(* IEC 61131-3 sources: 2026_Projet_YGO_ExcavatriceDragage/CODE/J_SUPERVISION/_TYPES/7_COMMUN_CONFIG, 11 files *)

(* ---- ST_BypassCommun.st ---- *)
(* ═══════════════════════════════════════════════════════════════
   ST_BypassCommun — Bypass maintenance GRANULAIRE, applicable aux 2 treuils à la fois
   ───────────────────────────────────────────────────────────────
   🎨 Distinct des bypass individuels M1/M2 (ST_BypassWinch)
      un OUI ici lève la protection sur LES DEUX treuils simultanément (pilotage "both",
      GVL_IHM.Commun.BtnWinchBothAscent/Descent), en OR avec le bypass individuel de chaque instance
      (PRG_04_Treuils_Benne). Évite de devoir activer 2 fois le même bypass (M1 ET M2) avant un
      pilotage groupé — SANS retirer les bypass individuels pour le pilotage à l'unité.
      ⚠️ Ne remplace PAS les bypass individuels : les deux se combinent en OR, jamais l'un
      n'entraîne la désactivation de l'autre.
   🔒 Doctrine : actionnable UNIQUEMENT en MAINT_N2, RETAIN, jamais masque
      les autres défauts du même bloc (voir REGISTRE_ACTIONS_Bypass_v1.0 (archive)).
   ═══════════════════════════════════════════════════════════════ *)
TYPE ST_BypassCommun :
STRUCT
    Global            : BOOL; (* 🌐 Bypass Global Commun (toutes sécurités communes M1+M2) *)
    SlackCable        : BOOL; (* ⚠️ Bypass capteur mou de câble — capteur unique M1/M2, OR avec bypass individuel *)
    TopLimitSwitch    : BOOL; (* 🚧 Bypass fin de course physique haute (capteur, bit5), OR avec bypass individuel *)
    TopLimitSoftware  : BOOL; (* : Bypass fin de course logiciel haut (position calculée), OR avec bypass individuel *)
    CableLimitSwitch  : BOOL; (* : Bypass limite basse physique (longueur câble), OR avec bypass individuel *)
    LimitLegal        : BOOL; (* : Bypass limite légale de profondeur, OR avec bypass individuel *)
    Initialized       : BOOL; (* Initialisé au boot *)
END_STRUCT
END_TYPE

(* ---- ST_BypassNetwork.st ---- *)
(* ═══════════════════════════════════════════════════════════════
   🌐 ST_BypassNetwork — Bypass général du diagnostic réseau
   ───────────────────────────────────────────────────────────────
   🔒 Permet de forcer les esclaves réseau (CAN, EtherCAT) à "online"
      pour le diagnostic, sans devoir toucher à chaque bit individuel.
      Jamais actif en production.
   ═══════════════════════════════════════════════════════════════ *)
TYPE ST_BypassNetwork :
STRUCT
    (* 📡 1. Bus maîtres & Modules d'E/S *)
    BusCanOpen  : BOOL; (* 📡 Bypass diagnostic bus CANopen maître *)
    BusEthercat : BOOL; (* 📡 Bypass diagnostic bus EtherCAT maître *)
    InputModules: BOOL; (* 🩺 Bypass diagnostic des 5 modules d'E/S physiques *)

    (* 🕹️ 2. Équipements esclaves *)
    Joystick    : BOOL; (* 🕹️ Bypass diagnostic esclave CANopen Joystick *)
    EncoderM1   : BOOL; (* 🧲 Bypass diagnostic esclave EtherCAT COD1 (M1 codeur) *)
    EncoderM2   : BOOL; (* 🧲 Bypass diagnostic esclave EtherCAT COD2 (M2 codeur) *)
    VariateurM3 : BOOL; (* ↔️ Bypass diagnostic esclave EtherCAT AC600 (M3 drive) *)
    IhmHeartbeat: BOOL := TRUE; (* 💓 Bypass du bit de vie IHM (défaut TRUE = sécurisé si pas d'IHM) *)

    (* 🛡️ 3. Hiérarchie & Restauration *)
    Global      : BOOL; (* 🌐 Bypass Global : tous les bus et esclaves réseau à la fois *)
    // Flag restauration boot dédié (défaut FALSE non ambigu, contrairement à une valeur métier)
    Initialized : BOOL := FALSE; (* 🚦 TRUE = bypass restauré depuis GVL_BypassRetain ce boot *)
END_STRUCT
END_TYPE

(* ---- ST_BypassSync.st ---- *)
(* ═══════════════════════════════════════════════════════════════
   ST_BypassSync — Bypass de la surveillance synchronisation M1/M2
   🔒 Doctrine : actionnable UNIQUEMENT en MAINT_N2, RETAIN, jamais masque
      les autres défauts du même bloc (voir REGISTRE_ACTIONS_Bypass_v1.0 (archive)).
   ═══════════════════════════════════════════════════════════════ *)
TYPE ST_BypassSync :
STRUCT
    Global      : BOOL := FALSE; (* 🌐 Bypass GLOBAL synchro : ignore toute erreur de synchronisation *)
    Initialized : BOOL := FALSE; (* 🚦 flag restauration boot *)
END_STRUCT
END_TYPE

(* ---- ST_CommunCfg.st ---- *)
(* ═══════════════════════════════════════════════════════════════
   ST_CommunCfg — Configuration des paramètres communs machine
   ═══════════════════════════════════════════════════════════════ *)
TYPE ST_CommunCfg :
STRUCT
    // Blocage instantané à 0m : sans défaut explicite,
    // ce champ vaut 0.0 tant qu'il n'a pas été réglé côté IHM -- "CablePosM <= 0.0" se déclenche
    // dès la position de référence, avant tout réglage réel de la cote légale. Défaut -999.0
    // (jamais atteint en pratique) : LimitLegalEnabled=TRUE sans réglage ne bloque plus rien par
    // erreur -- il faut régler la vraie cote pour que la protection devienne active.
    LimitLegalDepthMinAllowed_M : REAL := -30.0; (* 📐 Cote min de dragage autorisée (m, négatif) *)
    LimitLegalEnabled           : BOOL; (* 🟢 Activation de la limite légale *)
    SelHomingApproachEnable     : BOOL; (* 🔌 Case IHM : autorise le dépassement butée haute pour homing (si MAINT_N2) *)
    WinchMaxStepDescent      : INT := 5;     (* 🚀 Plafond palier descente nominal (1..5), commun M1/M2 *)
    WinchMaxStepAscent          : INT := 5;     (* 🚀 Limitation palier vitesse en montée (1..5), commun M1/M2 *)
    WinchSlowdownDistanceTop_M     : REAL := 0.5;  (* 📏 Distance avant limite haute : 0 = arrêt au seuil (m), commun M1/M2 *)
    WinchSlowdownDistanceBottom_M  : REAL := 1.0;  (* 📏 Distance avant limite basse pour ralentir (m), commun M1/M2 *)
    // : WinchSlowSpeed_Pct (%) retiré — un treuil ne connaît que des paliers (1..5),
    // pas une vitesse continue.
    WinchSlowdownMaxStep        : INT := 1;     (* : Plafond palier dans la zone de ralentissement (1..5), commun M1/M2 *)
    CfgCableLimitAscent_M       : REAL := 7.5;  (* 📐 Limite haute d'exploitation NORMALE (m), commun M1/M2 *)
    TglEnableKoboldAutoStopDescent : BOOL := FALSE; (* : Arrêt auto descente sur détection fond Kobold (pilotage normal) *)
    // Séquencement auto benne en pilotage couplé (WinchSel=0, MAINT_N1/N2) :
    // pousser le joystick benne pas ouverte -> ouvre d'abord puis descend couplé ;
    // tirer benne pas fermée -> ferme d'abord puis remonte couplé.
    // Défaut TRUE (activé) ; 1 bouton IHM pour désactiver -> comportement brut
    // (2 treuils sans condition). OFF = jamais gouverné par instBucket.Busy hors
    // action MANUELLE benne (WinchSel=2) / DumpAtTremie / ExtractionAssist.
    TglEnableCoupledBucketSequencing : BOOL := TRUE;
    // 🔒 Verrouillage descente treuil M1/M2 en mode MAINT si le pont M3 n'est pas à P1/Maintenance :
    // Défaut TRUE (sécurisé) ; bouton IHM pour désactiver (permet descente treuils partout).
    TglEnableWinchDescentLock_M3 : BOOL := TRUE;
    Initialized                 : BOOL := FALSE; (* 🚦 flag restauration boot *)
END_STRUCT
END_TYPE

(* ---- ST_CommunHMI.st ---- *)
(* ═══════════════════════════════════════════════════════════════
   🌐 ST_CommunHMI — Données d'échange IHM COMMUNES (pas propres à un axe)
   ───────────────────────────────────────────────────────────────
   Regroupe les signaux qui ne concernent
   PAS un axe/mécanisme en particulier (1 seul capteur/signal partagé par toute la
   machine) — évite de les dupliquer ou de les laisser en variables isolées
   directement dans GVL_IHM. Exemple : TopPositionSensorActive (capteur unique,
   commun M1+M2), BrakeThermalFault (retour unique, commun M1+M2+M3).
   ⚠️ Ne pas y mettre HmiInitDone (indicateur interne de séquencement boot, pas une
   information machine destinée à l'opérateur) — reste seul dans GVL_IHM.
   🧭 Structuration homogène : états → Cfg → Bypass (Cfg au-dessus de Bypass,
   Bypass en bas), cohérent avec ST_WinchHMI / ST_SyncHMI.
   ═══════════════════════════════════════════════════════════════ *)
TYPE ST_CommunHMI :
STRUCT
    TopPositionSensorActive   : BOOL; (* ⚠️ Capteur de position haute commun M1+M2 détecté *)
    TopHardStopLatched        : BOOL; (* 🔒 Latch directionnel capteur position haute commun M1+M2 actif *)
    BrakeThermalFault         : BOOL; (* 🌡️ Défaut/perte thermique frein — retour unique commun M1/M2/M3, escalade PowerCutOff *)
    PhaseRotationFault        : BOOL; (* ⚡ Rotation de phase incorrecte — retour unique commun M1/M2/M3
                                          (auparavant invisible IHM, seulement décodable via SafetyErrorId bit4/bit2) *)
    LimitLegalReached         : BOOL; (* 📐 Limite légale de profondeur de dragage atteinte (globale) *)
    HydraulicThermalFault     : BOOL; (* 🌡️ Défaut/perte thermique centrale hydraulique
                                          (PRG_02_Acquisition, diagnostic seul — aucune commande PLC) *)

    (* 🩺 Indicateurs diagnostic bypass — PLC→IHM, état réellement consommé *)
    SimTopSensorBypassActive  : BOOL; (* 🩺 1 = Bypass.TopLimitSwitch réellement actif *)
    SimSlackCableBypassActive : BOOL; (* 🩺 1 = Bypass.SlackCable réellement actif *)
    WinchInputSourceChanged   : BOOL; (* 🔀 PLC→IHM : source Winch a basculé (réel/simu) ce cycle *)

    (* 💓 Heartbeat IHM↔PLC — IHM inverse TglHeartbeatIhm toutes les 500 ms. *)
    TglHeartbeatIhm        : BOOL; (* IHM→PLC : toggle périodique, jamais valeur constante *)
    TglHeartbeatPlc        : BOOL; (* PLC→IHM : clignotant activité PLC *)
    HeartbeatIhmOk            : BOOL; (* PLC→IHM : front IHM post-boot reçu et timeout absent *)
    HeartbeatIhmTimeout       : BOOL; (* PLC→IHM : aucun front IHM depuis 2 s *)
    HeartbeatIhmElapsed       : TIME; (* PLC→IHM : temps depuis dernier front IHM *)

    // Boutons pilotage direct des 2 treuils (communs, remplace SelJoystickWinch en mode boutons)
    BtnWinchBothAscent     : BOOL; (* ⬆️ Monte les 2 treuils simultanément *)
    BtnWinchBothDescent   : BOOL; (* ⬇️ Descend les 2 treuils simultanément *)

    // Alarme restauration config PERSISTENT (RETAIN invalidé, ex. changement de
    // struct ST_*HMI) — visible et acquittable, jamais de disparition automatique silencieuse
    // (doctrine reset=front, PRG_07_Supervision.st §2bis). Vérifier les valeurs avant reprise cycle.
    ConfigRestoredFromPersistent : BOOL; (* ⚠️ PLC→IHM : restauration détectée ce boot, à vérifier *)
    BtnAckConfigRestored         : BOOL; (* 🔘 IHM→PLC : acquittement opérateur (front) *)

    Preflight : ST_PreflightHMI; (* 🩺 Verdict observateur à l'arrêt — jamais bloquant *)
    WinchSymmetry : ST_WinchSymmetryHMI; (* ⚖️ Mesures passives M1/M2 *)

    (* 🩺 Diagnostic arrêt auto descente Kobold (pilotage normal) *)
    KoboldImmersionConfirmed : BOOL; (* Front Kobold confirmé dans la fenêtre d'immersion *)
    KoboldBottomTouchLatched : BOOL; (* Fond détecté, descente bloquée (ProcessPermitM1/M2_Descend) *)

    (* ⏱️ Compteurs horaires maintenance — Machine (PLC sous tension) + M1/M2/M3 (marche reelle) *)
    RunningHours : ST_RunningHoursHMI;

    (* ⚙️ Configuration technologique codeur commune M1/M2 *)
    EncoderCfg : ST_fbEncoder_Cfg; (* Réglage mode confirmation preset, ponté vers GVL_PERSISTENT *)

    (* 📐 Configuration des paramètres communs machine (au-dessus des bypass) *)
    Cfg : ST_CommunCfg;

    (* 🔒 Bypass maintenance de capteurs COMMUNS (voir REGISTRE_ACTIONS_Bypass_v1.0 (archive)) *)
    Bypass : ST_BypassCommun;    (* 🔒 Granulaire, applique le bypass aux 2 treuils simultanément (pilotage "both") — OR avec le bypass individuel M1/M2 dans PRG_04 *)
END_STRUCT
END_TYPE

(* ---- ST_LocalIHM.st ---- *)
(* =======================================================================
   ST_LocalIHM — Échange cyclique IHM local
   -----------------------------------------------------------------------
   📄 Frontière : GVL_IHM.LocalIHM
   🎯 Rôle : regrouper les blocs de commandes et d'états de l'IHM locale.
   ======================================================================= *)
TYPE ST_LocalIHM :
STRUCT
    CtrlBlock   : ST_LocalIHM_CtrlBlock;   // IHM→PLC : commandes cycliques locales
    StatusBlock : ST_LocalIHM_StatusBlock; // PLC→IHM : états cycliques locaux
END_STRUCT
END_TYPE

(* ---- ST_RunningHoursHMI.st ---- *)
(* ═══════════════════════════════════════════════════════════════
   ⏱️ ST_RunningHoursHMI — Compteurs horaires maintenance (PLC→IHM)
   ───────────────────────────────────────────────────────────────
   🎯 Role : totalisateurs de marche pour planification maintenance,
      independants du chrono de cycle (qui se remet a zero par passe).
   🔌 Machine = duree sous tension PLC (toujours active des le boot).
      M1/M2/M3 = duree contacteur marche reel actif (preuve physique).
   💾 Source RETAIN : GVL_PERSISTENT (secondes), converties ici en H:Min.
   ═══════════════════════════════════════════════════════════════ *)
TYPE ST_RunningHoursHMI :
STRUCT
    MachineHours_H   : DINT; (* Heures entieres, PLC sous tension *)
    MachineHours_Min : INT;  (* Minutes 0..59 *)
    M1Hours_H        : DINT; (* Heures entieres, treuil M1 en marche *)
    M1Hours_Min      : INT;
    M2Hours_H        : DINT; (* Heures entieres, treuil M2 en marche *)
    M2Hours_Min      : INT;
    M3Hours_H        : DINT; (* Heures entieres, translation M3 en marche *)
    M3Hours_Min      : INT;
END_STRUCT
END_TYPE

(* ---- ST_SyncCfg.st ---- *)
(* ═══════════════════════════════════════════════════════════════
   ST_SyncCfg — Configuration de la synchronisation M1/M2
   ═══════════════════════════════════════════════════════════════ *)
TYPE ST_SyncCfg :
STRUCT
    CfgSyncTolerance_M : REAL := 3.0;   (* 📐 Tolérance max d'écart (m) — Dégradation Palier 1 dès 3.0m *)
    CfgSyncCriticalTolerance_M : REAL := 6.0; (* 🔴 Seuil 2 critique (m) — blocage synchro ; doit être > CfgSyncTolerance_M *)
    Initialized        : BOOL := FALSE; (* 🚦 Flag restauration boot (config restaurée depuis GVL_PERSISTENT) *)
END_STRUCT
END_TYPE

(* ---- ST_SyncCmd.st ---- *)
(* ═══════════════════════════════════════════════════════════════
   🎮 ST_SyncCmd — Commandes IHM pour la synchronisation M1/M2
   ═══════════════════════════════════════════════════════════════ *)
TYPE ST_SyncCmd :
STRUCT
    SelSyncEnable : BOOL := TRUE; (* ☑️ coché = synchro voulue (MAINT_N1/N2) *)
END_STRUCT
END_TYPE

(* ---- ST_SyncHMI.st ---- *)
(* ═══════════════════════════════════════════════════════════════
   ⚙️ ST_SyncHMI — Données d'échange IHM pour la synchronisation M1/M2
   ───────────────────────────────────────────────────────────────
   📄 Structuration en Cmd / State / Cfg / Bypass , homogène avec ST_WinchHMI.
   ═══════════════════════════════════════════════════════════════ *)
TYPE ST_SyncHMI :
STRUCT
    Cmd    : ST_SyncCmd;
    State  : ST_SyncState;
    Cfg    : ST_SyncCfg;
    Bypass : ST_BypassSync;
END_STRUCT
END_TYPE

(* ---- ST_SyncState.st ---- *)
(* ═══════════════════════════════════════════════════════════════
   🚦 ST_SyncState — États et diagnostics de la synchronisation M1/M2
   ═══════════════════════════════════════════════════════════════ *)
TYPE ST_SyncState :
STRUCT
    DeltaPos_M : REAL;    (* 📊 Écart de position réel mesuré (m) *)
    SyncActive : BOOL;    (* ⚖️ Indicateur si surveillance active *)
    SyncWarn   : BOOL;    (* ⚠️ LED d'alarme écart hors tolérance *)
    SyncDeviationWarn : BOOL; (* 🐢 Écart modéré actif : limitation forcée au Palier 1 *)
    Ready      : BOOL;    (* 🟢 Bloc de synchro prêt *)
    Error        : BOOL;    (* Alarme synchro active *)
    FaultLatched : BOOL;    (* 🔒 Défaut synchro latché (acquittable Reset) *)
    ErrorId      : WORD;    (* ❌ Code défaut synchro *)
    FBState    : E_State; (* 🤖 État de l'automate interne (FB_WinchSync) *)
END_STRUCT
END_TYPE
